TYPE U_YARD_CTRL :
UNION
  stCtrl              : ST_YARD_CTRL;
  byCtrl    AT %Q*    : ARRAY[1..SIZEOF(ST_YARD_CTRL)] OF BYTE;
END_UNION
END_TYPE

(* stored: Version 1.1.0.1
   DUT U_YARD_CTRL: Id {1de2f777-4d3b-49ff-be8d-d327c3f3e543} *)
